// TIA Portal V20 export
// export: Created 2026-10-19T18:37:16.7483408Z, ExportSetting WithDefaults, DisplayName Totally Integrated Automation Portal, DisplayVersion V20 Update 6, DisplayName TIA Portal Openness, DisplayVersion V20 Update 6, DisplayName TIA Portal Version Control Interface, DisplayVersion V20 Update 6, DisplayName SINAMICS Startdrive Advanced, DisplayVersion V20 SP1, DisplayName SINAMICS Startdrive G130, G150, S120, S150, SINAMICS MV, G220, S200, S210, DisplayVersion V20 SP1, DisplayName SINAMICS Startdrive G110M, G120, G120C, G120D, G120P, G115D, DisplayVersion V20 SP1, DisplayName STEP 7 Professional, DisplayVersion V20 Update 6, DisplayName STEP 7 Safety, DisplayVersion V20 Update 2, DisplayName WinCC Basic/Comfort/Advanced, DisplayVersion V20 Update 6, DisplayName WinCC Unified, DisplayVersion V20 Update 6
DATA_BLOCK "OrderTable_HMI"   // DB96
{ S7_Optimized_Access := 'TRUE' }
VERSION : 0.1
// stored: AutoNumber true, DBAccessibleFromOPCUA true, IsOnlyStoredInLoadMemory false, IsRetainMemResEnabled false, IsWriteProtectedInAS false, MemoryReserve 100
   VAR
      Start : Bool;
      Pause : Bool;
      Resume : Bool;
      Stop : Bool;
      "Manual order" : Bool;
      Transfer_From_To : Byte;
      "Send VTD Order" : Bool;
      "Send CNV Order" : Bool;
      "From level" : Byte;
      "To level" : Byte;
      "Testing Time" : UInt;
      "Numer of cycles" : Byte;
      Level : Byte;
      "Time Running" : UInt;
      Actual_Cycle : Byte;
      "Start Test Visibility" : Bool;
      "Stop Test Visibility" : Bool;
      "Pause Test Visibility" : Bool;
      "Resume Visibility" : Bool;
      "Clear Table Visibility" : Bool;
      Auto_Settings_Visibility : Bool;
      "Manual order Visibility" : Bool;
      "VTD_Manual_Orders Visibility" : Bool;
      "Buffers_Manual_Orders Visibility" : Bool;
      "Send VTD Order Visibility" : Bool;
      "Send CNV Order Visibility" : Bool;
      Transfer_CNV1_L6 : Bool;
      Transfer_CNV1_L5 : Bool;
      Transfer_CNV1_L4 : Bool;
      Transfer_CNV1_L3 : Bool;
      Transfer_CNV1_L2 : Bool;
      Transfer_CNV2_L6 : Bool;
      Transfer_CNV2_L5 : Bool;
      Transfer_CNV2_L4 : Bool;
      Transfer_CNV2_L3 : Bool;
      Transfer_CNV2_L2 : Bool;
      Transfer_Out_VTD : Bool;
      Transfer_Into_VTD : Bool;
      Occupied_CNV1_L6 : Bool;
      Occupied_CNV1_L5 : Bool;
      Occupied_CNV1_L4 : Bool;
      Occupied_CNV1_L3 : Bool;
      Occupied_CNV1_L2 : Bool;
      Occupied_CNV2_L6 : Bool;
      Occupied_CNV2_L5 : Bool;
      Occupied_CNV2_L4 : Bool;
      Occupied_CNV2_L3 : Bool;
      Occupied_CNV2_L2 : Bool;
      Occupied_Buffer_VTD : Bool;
      Occupied_Extractor_VTD : Bool;
      CurrentLevel : UInt;
   END_VAR
BEGIN
END_DATA_BLOCK
